FUNCTION_BLOCK FB_Runtime_Test EXTENDS TcUnit.FB_TestSuite
VAR_INPUT
END_VAR
VAR_OUTPUT
END_VAR
VAR
END_VAR

elapsedTimeShouldBe5sAfter5s();
elapsedFlagShouldBeTrueAfterSettimePassed();
elapsedFlagShouldntBeTrueBeforeSettimePassed();
elapsedTimeShouldBe7seconds();
elapsedTimeShouldBeLessThanStartTimeWhenCountdownUsed();

METHOD elapsedFlagShouldBeTrueAfterSettimePassed
VAR
	runtime : FB_Runtime;
END_VAR

TEST('elapsedFlagShouldBeTrueAfterSettimePassed');

	runtime.setTestMode(
		testtime := T#5S,
		reset := FALSE);

	runtime(
		gotime:= TRUE, 
		settime:= T#5S, 
		countdown:= , 
		resetToTime:= , 
		elapsedtime=> , 
		elapsed=> );
		
	runtime(
		gotime:= TRUE, 
		settime:= T#5S, 
		countdown:= , 
		resetToTime:= , 
		elapsedtime=> , 
		elapsed=> );

	AssertEquals_BOOL(Expected :=  TRUE, Actual := runtime.elapsed , Message := 'Elapsed flag not true after settime passed');	

TEST_FINISHED();
END_METHOD

METHOD elapsedFlagShouldntBeTrueBeforeSettimePassed
VAR
	runtime : FB_Runtime;
END_VAR

TEST('elapsedFlagShouldntBeTrueBeforeSettimePassed');

	runtime.setTestMode(
		testtime := T#4900MS,
		reset := FALSE);

	runtime(
		gotime:= TRUE, 
		settime:= T#5S, 
		countdown:= , 
		resetToTime:= , 
		elapsedtime=> , 
		elapsed=> );


	AssertEquals_BOOL(Expected :=  FALSE, Actual := runtime.elapsed , Message := 'Elapsed flag not false before settime passed');	

TEST_FINISHED();
END_METHOD

METHOD elapsedTimeShouldBe5sAfter5s : BOOL
VAR
	runtime : FB_Runtime;
END_VAR

TEST('elapsedTimeShouldBe5sAfter5ss');

	runtime.setTestMode(
		testtime := T#4990MS,
		reset := FALSE);

	runtime(
		gotime:= TRUE, 
		settime:= T#10S, 
		countdown:= , 
		resetToTime:= , 
		elapsedtime=> , 
		elapsed=> );

	AssertEquals_BOOL(Expected :=  TRUE, Actual := runtime.elapsedTime = T#5S , Message := 'Elapsed time not 5s after 5s!');	

TEST_FINISHED();
END_METHOD

METHOD elapsedTimeShouldBe7seconds
VAR
	runtime : FB_Runtime;
END_VAR

TEST('elapsedTimeShouldBe7seconds');

	runtime.setTestMode(
		testtime := T#7010MS,
		reset := FALSE);

	runtime(
		gotime:= FALSE, 
		settime:= T#10S, 
		countdown:= TRUE, 
		resetToTime:= , 
		elapsedtime=> , 
		elapsed=> );

	AssertEquals_BOOL(Expected :=  TRUE, Actual := runtime.elapsedTime = T#7S , Message := 'Elapsed time not 7s!');	

TEST_FINISHED();
END_METHOD

METHOD elapsedTimeShouldBeLessThanStartTimeWhenCountdownUsed
VAR
	runtime : FB_Runtime;
END_VAR

TEST('elapsedTimeShouldBeLessThanStartTimeWhenCountdownUsed');

	runtime.setTestMode(
		testtime := T#7S,
		reset := FALSE);

	runtime(
		gotime:= FALSE, 
		settime:= T#10S, 
		countdown:= TRUE, 
		resetToTime:= , 
		elapsedtime=> , 
		elapsed=> );
		
	runtime(
		gotime:= FALSE, 
		settime:= T#10S, 
		countdown:= TRUE, 
		resetToTime:= , 
		elapsedtime=> , 
		elapsed=> );
		
	runtime(
		gotime:= FALSE, 
		settime:= T#10S, 
		countdown:= TRUE, 
		resetToTime:= , 
		elapsedtime=> , 
		elapsed=> );

	AssertEquals_BOOL(Expected :=  TRUE, Actual := runtime.elapsedTime < T#7S , Message := 'Elapsed time not less than start time when countdown used');	

TEST_FINISHED();
END_METHOD

END_FUNCTION_BLOCK

(* stored: Version 1.1.0.1, ProductVersion 3.1.4024.9
   POU FB_Runtime_Test: Id {a8d3d2e6-1af7-4f13-b66b-339c27657ac2}, SpecialFunc None
   Method elapsedFlagShouldBeTrueAfterSettimePassed: Id {c550d865-167f-49c2-a36b-3d2fe2643690}
   Method elapsedFlagShouldntBeTrueBeforeSettimePassed: Id {6c443bf9-7c32-4e14-876d-5004a00adc8d}
   Method elapsedTimeShouldBe5sAfter5s: Id {5972ffc9-b360-4674-a0ca-d70041eda663}
   Method elapsedTimeShouldBe7seconds: Id {c6a651f3-694a-4e66-aa7c-48e7b312ab8a}
   Method elapsedTimeShouldBeLessThanStartTimeWhenCountdownUsed: Id {4c8841b3-4a43-4dc4-8951-bb0a0795af18} *)
